// TIA Portal V21 export
// export: Created 2026-11-21T16:00:28.7892337Z, ExportSetting WithDefaults, DisplayName Totally Integrated Automation Portal, DisplayVersion V21, DisplayName STEP 7 Professional, DisplayVersion V21, DisplayName STEP 7 Safety, DisplayVersion V21, DisplayName Tech WebApplication, DisplayVersion V21, DisplayName WinCC Basic/Comfort/Advanced, DisplayVersion V21, DisplayName WinCC Unified, DisplayVersion V21
VAR_GLOBAL   // PLC tag table "Dosing"
   Dose_Level AT %IW64 : Int;   // Level of the dosing tank in percent
   Dose_Speed AT %MW10 : Int;   // Speed of the dosing pump
   Dose_Target AT %MW12 : Int;   // Target level
   Dose_Valve AT %Q0.0 : Bool;   // The dosing valve is open
END_VAR
